Fanuc KAREL source: kf00038.KL

-- PROVISIONAL review KL for V1013-1; original PC SHA256 dd93c658b368dab79bbf8d4661bd35aaf3a7a4c60de58a6ac1a81db5f768aa20
-- Incomplete behavior may be omitted. Consult companion uncertainty JSON. Do not deploy.
PROGRAM KF00038
%NOLOCKGROUP
VAR
  I : INTEGER
  J : INTEGER
  X : REAL
  Y : REAL
  B : BOOLEAN
  C : BOOLEAN
  TXT : STRING[80]
  TXT2 : STRING[80]
  STATUS : INTEGER
-- UNRESOLVED_DECL AI type=002010
-- UNRESOLVED_DECL BI type=002010
-- UNRESOLVED_DECL P type=000102
-- UNRESOLVED_DECL JP type=000199
-- UNRESOLVED_DECL PF type=000101
-- UNRESOLVED_DECL V1 type=000013
-- UNRESOLVED_DECL V2 type=000013
BEGIN
  -- UNRESOLVED_PC offsets 5-19; opcodes 2E,22,9D,33,35
  -- UNRESOLVED_PC offsets 24-38; opcodes 22,22,1E
  -- UNRESOLVED_PC offsets 43-47; opcodes 7F
END KF00038
